// TIA Portal V20 export
ORGANIZATION_BLOCK "Startup"   // OB100, LAD, Startup
TITLE = Startup
{ S7_Optimized_Access := 'TRUE' }
AUTHOR : IA
FAMILY : PRUEBA
VERSION : 0.1
// Tanda 7: Startup, incrementa Arranques
// stored: AutoNumber false, IsIECCheckEnabled false, SetENOAutomatically false
   VAR_INPUT
      LostRetentive : Bool;
      LostRTC : Bool;
   END_VAR
BEGIN

REGION Network 1: Contador de vida
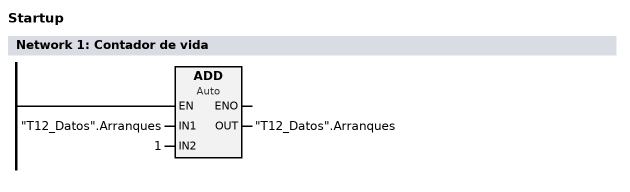
   RUNG wire#powerrail
      Add(in1 := "T12_Datos".Arranques, in2 := 1, out => "T12_Datos".Arranques)
   END_RUNG
   // the same network as SCL:
   "T12_Datos".Arranques := "T12_Datos".Arranques + 1;
END_REGION
END_ORGANIZATION_BLOCK
